(* IEC 61131-3 sources: PortalRobot/Portal_robot/Device/application/ST/ST_ROBOT, 16 files *)

(* ---- E_ROBOT_ACTION.st ---- *)
{attribute 'qualified_only'}
{attribute 'strict'}
TYPE E_ROBOT_ACTION :
(
	NONE,
	MOVE_TO_POINT,
	UNCLAMP_1,
	CLAMP_1,
	UNCLAMP_2,
	CLAMP_2,
	ROTATE_TO_BLANK,
	ROTATE_TO_DETAIL

);
END_TYPE

(* ---- E_ROBOT_CONTROL_MODE.st ---- *)
{attribute 'qualified_only'}
{attribute 'strict'}
TYPE E_ROBOT_CONTROL_MODE :
(
	SOFTMOTION := 0,
	MODBUS_TCP := 1
);
END_TYPE

(* ---- E_ROBOT_MODBUS_CLIENT_STATE.st ---- *)
{attribute 'qualified_only'}
{attribute 'strict'}
TYPE E_ROBOT_MODBUS_CLIENT_STATE :
(
	DISABLED,
	CONNECTING,
	INITIAL_READ,
	INITIAL_READ_RELEASE,
	CLEAR_COMMAND,
	CLEAR_COMMAND_RELEASE,
	READY,
	WRITE_COMMAND,
	WRITE_COMMAND_RELEASE,
	READ_STATUS,
	READ_STATUS_RELEASE,
	RECONNECT_WAIT
);
END_TYPE

(* ---- E_ROBOT_MODBUS_EXECUTION_STATE.st ---- *)
{attribute 'qualified_only'}
{attribute 'strict'}
TYPE E_ROBOT_MODBUS_EXECUTION_STATE :
(
	IDLE := 0,
	ACCEPTED := 1,
	BUSY := 2,
	DONE := 3,
	ERROR := 4,
	STOPPED := 5
);
END_TYPE

(* ---- E_ROBOT_STATE.st ---- *)
{attribute 'qualified_only'}
{attribute 'strict'}
TYPE E_ROBOT_STATE :
(
	IDLE,
	MOTION,
	GRIPPER,
	DONE,
    ERROR,
	MODBUS
);
END_TYPE

(* ---- ST_ROBOT_COMMAND.st ---- *)
TYPE ST_ROBOT_COMMAND :
STRUCT
	xExecute : BOOL; // Команда запуска
	xStop    : BOOL; // Команда остановки
	xReset   : BOOL; // Команда сброса внешнего робота
	eAction  : E_ROBOT_ACTION; // Элементарное действие робота
	eSetPoint: E_POINT_NAME; // Имя элементарной точки движения
	iActiveSlot : SINT; // Единственный слот, относительно которого выполняется команда
	uiMagazineId : UINT; // 0 вне магазина; 1 или 2 для точки соответствующего магазина
END_STRUCT
END_TYPE

(* ---- ST_ROBOT_DIAG.st ---- *)
TYPE ST_ROBOT_DIAG :
STRUCT
	eState        : E_ROBOT_STATE; // Текущее состояние автомата робота
	eActiveAction : E_ROBOT_ACTION; // Выполняемое действие робота
	eActivePoint  : E_POINT_NAME; // Целевая точка текущего движения
	stWarning     : ST_WARNING_EVENT; // Последнее предупреждение робота
END_STRUCT
END_TYPE

(* ---- ST_ROBOT_ERROR.st ---- *)
TYPE ST_ROBOT_ERROR :
STRUCT
	WRONG_ACTION : BOOL; // Получена неизвестная команда робота
	MOTION_ERROR : BOOL; // Ошибка менеджера движения
	GRIPPER_ERROR: BOOL; // Ошибка механизма захвата
	MODBUS_ERROR : BOOL; // Совместимость: любая ошибка внешнего интерфейса
	MODBUS_COMMUNICATION_ERROR : BOOL; // Ошибка TCP/FC03/FC16/heartbeat
	EXTERNAL_ROBOT_ALARM : BOOL; // Контроллер робота сообщил технологическую аварию
	STOP_ERROR   : BOOL; // Движение остановлено командой или глобальной ошибкой
END_STRUCT
END_TYPE

(* ---- ST_ROBOT_ERRORS.st ---- *)
TYPE ST_ROBOT_ERRORS :
STRUCT
	dwErrorActive : DWORD; // Битовая маска активных ошибок
	dwErrorLast   : DWORD; // Битовая маска последних ошибок
	dwAlarmActive : DWORD; // Собственные аварии робота для общего журнала
	stErrorActive : ST_ROBOT_ERROR; // Расшифровка активных ошибок
	stErrorLast   : ST_ROBOT_ERROR; // Расшифровка последних ошибок
END_STRUCT
END_TYPE

(* ---- ST_ROBOT_FAULT_REQUEST.st ---- *)
TYPE ST_ROBOT_FAULT_REQUEST :
STRUCT
	xEnabled     : BOOL; // Глобальное разрешение диагностической инъекции
	xWrongAction : BOOL; // Импульс недопустимого действия робота
	stGripper : ST_GRIPPER_FAULT_REQUEST; // Неисправности виртуального захвата
	stPoint   : ST_POINT_FAULT_REQUEST; // Ошибки проверки точки движения
END_STRUCT
END_TYPE

(* ---- ST_ROBOT_FAULT_STATUS.st ---- *)
TYPE ST_ROBOT_FAULT_STATUS :
STRUCT
	stRobot   : ST_FAULT_INJECTION_STATUS; // Локальная ошибка автомата робота
	stGripper : ST_FAULT_INJECTION_STATUS; // Неисправности виртуального захвата
	stPoint   : ST_FAULT_INJECTION_STATUS; // Ошибки проверки точки движения
END_STRUCT
END_TYPE

(* ---- ST_ROBOT_MODBUS_CONFIG.st ---- *)
TYPE ST_ROBOT_MODBUS_CONFIG :
STRUCT
	aIpAddress        : ARRAY [0..3] OF BYTE; // IPv4 контроллера робота
	uiPort            : UINT := UINT#502; // TCP-порт Modbus
	uiUnitId          : UINT := UINT#1; // Unit ID в Modbus TCP
	tResponseTimeout  : TIME := T#500MS; // Ожидание ответа FC03/FC16
	tPollInterval     : TIME := T#50MS; // Период чтения обратной связи
	tHeartbeatTimeout : TIME := T#2S; // Максимальная пауза heartbeat робота
	tCommandTimeout   : TIME := T#600S; // Предельная длительность одной команды
END_STRUCT
END_TYPE

(* ---- ST_ROBOT_MODBUS_STATUS.st ---- *)
TYPE ST_ROBOT_MODBUS_STATUS :
STRUCT
	xConfigValid       : BOOL; // Параметры соединения прошли проверку PLC
	xConnected         : BOOL; // TCP-соединение установлено
	xCommunicationAlive: BOOL; // Получена свежая обратная связь и меняется heartbeat
	xStatusFresh       : BOOL; // После подключения успешно прочитан блок 1101..1117
	xControllerOn      : BOOL;
	xAutomaticMode     : BOOL;
	xRemoteEnabled     : BOOL;
	xDrivesEnabled     : BOOL;
	xHomed             : BOOL;
	xEmergencyStop     : BOOL;
	xRobotAlarm        : BOOL;
	xPositionValid     : BOOL;
	xSimulatorActive   : BOOL; // Бит 1108.9: подключён Python-симулятор, а не реальный SC-500
	xReady             : BOOL; // Итоговая готовность, пересчитанная PLC
	xBusy              : BOOL;
	xDone              : BOOL;
	xError             : BOOL; // Ошибка исполнения, робота или транспорта
	xCommandTimeout    : BOOL; // Робот не завершил принятую команду за лимит
	xResetBusy         : BOOL; // Передача Reset и подтверждение его снятия ещё выполняются
	xResetDone         : BOOL; // Reset подтверждён обратной связью и очищенной FC16
	xResetFailed       : BOOL; // Попытка сорвана/истекла; повтор только новым запросом
	uiAckSeq           : UINT;
	uiExecutionState   : UINT;
	uiResultCode       : UINT;
	uiActiveCommand    : UINT;
	uiCurrentPoint     : UINT;
	uiGripperStatus    : UINT;
	uiRobotHeartbeat   : UINT;
	uiStatusWord       : UINT;
	uiAlarmCode        : UINT;
	uiOperationPhase   : UINT;
	uiProtocolVersion  : UINT;
	lrActualX          : LREAL;
	lrActualY          : LREAL;
	lrActualZ          : LREAL;
	udiClientError     : UDINT;
	udiReadError       : UDINT;
	udiWriteError      : UDINT;
END_STRUCT
END_TYPE

(* ---- ST_ROBOT_RESET_DEPENDENCIES.st ---- *)
TYPE ST_ROBOT_RESET_DEPENDENCIES :
STRUCT
	// Внутренний PLC-контракт: биты 0..2 — станки, 3..4 — магазины,
	// 5..6 — ГК, 7..8 — механизмы двухпалетных магазинов.
	dwStopOwners : DWORD; // Владельцы текущего зависимого ROBOT_STOP
	dwLiveCauses : DWORD; // Непосредственные удерживаемые причины этих владельцев
	dwResetBusy : DWORD; // Выполняющийся аппаратный/асинхронный сброс владельца
END_STRUCT
END_TYPE

(* ---- ST_ROBOT_RESET_RECOVERY.st ---- *)
TYPE ST_ROBOT_RESET_RECOVERY :
STRUCT
	udiAttempt : UDINT; // Ненулевой номер принятой попытки; не является HMI-командой
	xActive : BOOL; // Попытка ещё выполняется в FB_ROBOT
	xDependenciesReady : BOOL; // Первичные Motion/захват/Modbus восстановлены; ERROR родителя ещё допустим
END_STRUCT
END_TYPE

(* ---- ST_ROBOT_STATUS.st ---- *)
TYPE ST_ROBOT_STATUS :
STRUCT
	xBusy             : BOOL; // Робот выполняет команду
	xDone             : BOOL; // Команда завершена
	xError            : BOOL; // Робот находится в ошибке
	xExternalError    : BOOL; // Робот остановлен ошибкой зависимого блока
	xPowerAllowed     : BOOL; // Кнопка включения или отключения приводов доступна
	xStopAllowed      : BOOL; // Кнопка контролируемой остановки доступна
	xResetAllowed     : BOOL; // Кнопка сброса ошибок робота и приводов доступна
	eCurrentPoint     : E_POINT_NAME; // Последняя достигнутая точка
	uiMagazineContext : UINT; // 0 вне рабочей зоны; 1..2 — магазин, в рабочей зоне которого находится робот
	xBlankAvailable   : BOOL; // В первом захвате находится заготовка
	xDetailAvailable  : BOOL; // Во втором захвате находится готовая деталь
	uiBlankPayloadType  : UINT; // Фактический тип заготовки, 0 — неизвестно
	uiDetailPayloadType : UINT; // Фактический тип детали, 0 — неизвестно
	xGripper1Open     : BOOL; // Первый захват открыт
	xGripper1Closed   : BOOL; // Первый захват закрыт
	xGripper2Open     : BOOL; // Второй захват открыт
	xGripper2Closed   : BOOL; // Второй захват закрыт
	xRotatedToBlank   : BOOL; // Захват повёрнут к заготовке
	xRotatedToDetail  : BOOL; // Захват повёрнут к готовой детали
END_STRUCT
END_TYPE
